Fanuc KAREL source: kt00494.KL

-- PROVISIONAL review KL for V1013-1; original PC SHA256 dbbeddfe92da2c47cba980b16a510a7c3ba61403dc52837e7cdb0d78ce8f573e
-- Incomplete behavior may be omitted. Consult companion uncertainty JSON. Do not deploy.
PROGRAM KT00494
%NOLOCKGROUP
-- UNRESOLVED_DECL P1 type=000102
-- UNRESOLVED_DECL P2 type=000101
-- UNRESOLVED_DECL OUT type=000101
BEGIN
  -- UNRESOLVED_PC offsets 5-20; opcodes 2E,22,32,35
  -- UNRESOLVED_PC offsets 25-54; opcodes 49,7E,49,60,4A
  -- UNRESOLVED_PC offsets 59-63; opcodes 7F
END KT00494
